(* PLC project TBEN_L5_PLC11.project, CODESYS CODESYS V3.5 SP21 Patch 1 *)
(* stored: creationDateTime 2026-11-07T15:34:51.9760141, modificationDateTime 2026-11-07T15:09:07.4034196 *)

// Kết quả 1 request ISDU master trả cho client
TYPE ST_IolResult :
STRUCT
    xError         : BOOL;
    eErrSource     : E_IolErrSource;
    dwPnioStatus   : DWORD;                                // STATUS RDREC/WRREC
    uiIolMasterErr : UINT;                                 // IOL_M_ErrorCode
    uiIolDevErr    : UINT;                                 // lỗi ISDU device 0x80xx
    uiLen          : UINT;                                 // số byte dữ liệu đọc về
    abData         : ARRAY[0..GVL_IolConst.uiMAX_DATA - 1] OF BYTE;
END_STRUCT
END_TYPE
